Fanuc KAREL source: KO00125.KL

PROGRAM KO00125
%NOLOCKGROUP
VAR
  A: ARRAY[2] OF SHORT
  B: ARRAY[2] OF BYTE
  OUT: INTEGER
BEGIN
  A[1] = 1
  B[1] = 2
  OUT = ATAN2(A[1], B[1])
END KO00125
